TYPE TcoAteqG6_Inputs_v_3_5_x :
STRUCT
	{attribute addProperty Name "<#Input module 1 (slot 1, 00h..3Fh)#>"}
	In1 AT %I* : ARRAY[0..63] OF BYTE;
	{attribute addProperty Name "<#Input module 2 (slot 2, 40h..7Fh)#>"}
	In2 AT %I* : ARRAY[0..63] OF BYTE;
	{attribute addProperty Name "<#Input module 3 (slot 3, 80h..BFh)#>"}
	In3 AT %I* : ARRAY[0..63] OF BYTE;
	{attribute addProperty Name "<#Input module 4 (slot 4, C0h..FFh)#>"}
	In4 AT %I* : ARRAY[0..63] OF BYTE;
END_STRUCT
END_TYPE

(* stored: Version 1.1.0.1, ProductVersion 3.1.4024.12
   DUT TcoAteqG6_Inputs_v_3_5_x: Id {8d019df1-8ed4-4129-a599-d4b0ad86cbba} *)
